(* IEC 61131-3 sources: trust-platform/examples/OSCAT/weather_station_conversion/non-oop/src, 3 files *)

(* ---- Configuration.st ---- *)
CONFIGURATION WeatherStationConversionClassicConfiguration
RESOURCE Cpu0 ON PLC
    TASK MainTask (INTERVAL := T#1s, PRIORITY := 1);
    PROGRAM Main WITH MainTask : Main;
END_RESOURCE
END_CONFIGURATION

(* ---- Main.st ---- *)
PROGRAM Main
VAR
    ConstantsReady : BOOL;
    WindMetersPerSecond : REAL := REAL#10.0;
    WindDegrees : INT := INT#90;
    BeaufortIndex : INT;
    WindDirection : STRING[3];
END_VAR

ConstantsReady := OSCAT_BASIC_Constants();
BeaufortIndex := MS_TO_BFT(MS := WindMetersPerSecond);
WindDirection := DEG_TO_DIR(DEG := WindDegrees, N := INT#4, L := INT#1);
END_PROGRAM

(* ---- Tests.st ---- *)
TEST_PROGRAM WeatherStationConversionClassicConvertsWindData
VAR
    ConstantsReady : BOOL;
END_VAR

ConstantsReady := OSCAT_BASIC_Constants();

ASSERT_TRUE(IN := ConstantsReady);
ASSERT_EQUAL(EXPECTED := MS_TO_BFT(MS := REAL#10.0), ACTUAL := MS_TO_BFT(MS := REAL#10.0));
ASSERT_EQUAL(EXPECTED := DEG_TO_DIR(DEG := INT#90, N := INT#4, L := INT#1), ACTUAL := DEG_TO_DIR(DEG := INT#90, N := INT#4, L := INT#1));
END_TEST_PROGRAM
